Fanuc KAREL source: kt00568.KL

-- PROVISIONAL review KL for V1013-1; original PC SHA256 a92afe680aad82af2b8477d01129232d9ec67b163db568a400f18fa47914cd81
-- Incomplete behavior may be omitted. Consult companion uncertainty JSON. Do not deploy.
PROGRAM KT00568
%NOLOCKGROUP
VAR
  R2 : REAL
-- UNRESOLVED_DECL V1 type=000013
-- UNRESOLVED_DECL OUT type=000013
BEGIN
  -- UNRESOLVED_PC offsets 5-20; opcodes 2E,22,32,35
  -- UNRESOLVED_PC offsets 25-36; opcodes 2E,23
  -- UNRESOLVED_PC offsets 41-63; opcodes 49,21,8E,4A
  -- UNRESOLVED_PC offsets 68-72; opcodes 7F
END KT00568
